(* CODESYS project filelogger.library
   DefaultNamespace: KOSTAL.AF2024.Core.FileLogger
   DocFormat: reStructuredText
   Description: Contains Functionalities to log strings to Filesystem with WSTRING content
   Author: Frank Dümpelmann
   Title: KOSTAL.AF2024.Core.FileLogger
   Version: 1.0.0.0
   Company: KOSTAL GmbH & Co.KG
   Placeholder: KOSTAL.AF2024.Core.FileLogger

Project tree, tasks and I/O mapping:
  libraries: KOSTAL.AF2024.Core.functionResponse, 1.0.0.0 (KOSTAL GmbH & Co.KG); KOSTAL.AF2024.Core.GetSystemTime, 1.0.0.0 (KOSTAL GmbH & Co.KG); KOSTAL.AF2024.Core.Process, 1.0.0.0 (KOSTAL GmbH & Co.KG); KOSTAL.AF2024.Core.Settings, 1.0.0.0 (KOSTAL GmbH & Co.KG); KOSTAL.AF2024.Core.StringTools, 1.0.0.0 (KOSTAL GmbH & Co.KG); KOSTAL.AF2024.Core.System, 1.0.0.0 (KOSTAL GmbH & Co.KG); Tc2_Standard, 3.3.3.0 (Beckhoff Automation GmbH); Tc2_System, 3.6.2.0 (Beckhoff Automation GmbH); Tc2_Utilities, 3.5.2.0 (Beckhoff Automation GmbH)
  DUT/
  POU/
    Interface/
      interface I_Logger: ePath, Extension, Path, Prefix, amsNedId_fileServer, delimiter, enabled, ID, maxLine, name, reset, StackCount, State, stepNumber, timeout, addLine
      interface I_Logger_Owner: ePath, Extension, Path, Prefix, amsNedId_fileServer, delimiter, enabled, maxLine, timeout, linkTimeSource, resetLogger, stepNumber
    function block FB_FileLogger [ST]: _a0_Ready, _a1_FileExist, _a2_Close, _a2_Open, _a2_Write, _Add_UTF16_LE_Header, _addLine, _control, _device, _formatWordToString, _getFqFileName, _outOfLimitControl, _stepHeader, _write, ePath, Extension, Path, Prefix, amsNedId_fileServer, delimiter, enabled, ID, maxLine, name, reset, StackCount, State, stepNumber, timeout, addLine, linkTimeSource, resetLogger, FBmain
  Project Information/
    function F_GetCompany [ST]
    function F_GetTitle [ST]
    function F_GetVersion [ST]
  Version/
    global variables Global_Version
*)

// Version/Global_Version
{attribute 'TcGenerated'}
{attribute 'no-analysis'}
{attribute 'linkalways'}
// This function has been automatically generated from the project information.
VAR_GLOBAL CONSTANT
	{attribute 'const_non_replaced'}
	stLibVersion_KOSTAL_AF2024_Core_FileLogger : ST_LibVersion := (iMajor := 1, iMinor := 0, iBuild := 0, iRevision := 0, nFlags := 0, sVersion := '1.0.0.0');
END_VAR

// POU/Interface/I_Logger
INTERFACE I_Logger EXTENDS KOSTAL_AF2024_Core_System.I_Interface

PROPERTY PUBLIC ePath : Tc2_System.E_OpenPath
GET
END_GET
END_PROPERTY

(*
Description
===========
| Extension of the saved file
| Default: .log
*)
PROPERTY PUBLIC Extension : STRING
GET
END_GET
END_PROPERTY

(*
Description
===========
| File path and name WITHOUT file extension
| e.g. "C:\\Logs\\test" creates the file "C:\\Logs\\test.log"
| default: c:\\temp\\log
*)
PROPERTY PUBLIC Path : KOSTAL_AF2024_Core_Settings.T_MaxString_UTF8
GET
END_GET
END_PROPERTY

PROPERTY PUBLIC Prefix : KOSTAL_AF2024_Core_Settings.T_MaxString_UTF8
GET
END_GET
END_PROPERTY

(*
Description
===========
| AMS NetID of  device to save log file to
| default: '' = Local device
*)
PROPERTY PUBLIC amsNedId_fileServer : STRING
GET
END_GET
END_PROPERTY

(*
Description
===========
| Delimiter to separate log records
| default: ;
*)
PROPERTY PUBLIC delimiter : WSTRING(1)
GET
END_GET
END_PROPERTY

(*
Description
===========
| Reset file handling sequence 
*)
PROPERTY PUBLIC enabled : BOOL
GET
END_GET
END_PROPERTY

PROPERTY ID : WSTRING
GET
END_GET
SET
END_SET
END_PROPERTY

(*
Description
===========
| Maximum number of message lines in write queue. 
| If the number is exceeded, the lines will be discarded
| default: 100, Maximum: 255
*)
PROPERTY PUBLIC maxLine : UDINT
GET
END_GET
END_PROPERTY

PROPERTY name : WSTRING
GET
END_GET
SET
END_SET
END_PROPERTY

(*
Description
===========
| Reset file handling sequence 
*)
PROPERTY PUBLIC reset : BOOL
GET
END_GET
END_PROPERTY

PROPERTY PUBLIC StackCount : UDINT
GET
END_GET
END_PROPERTY

PROPERTY PUBLIC State : KOSTAL_AF2024_Core_functionResponse.I_T_functionResponse
GET
END_GET
END_PROPERTY

PROPERTY stepNumber : INT
GET
END_GET
SET
END_SET
END_PROPERTY

(*
Description
===========
| Maximum time allowed for write operation
| default: 5s
*)
PROPERTY PUBLIC timeout : TIME
GET
END_GET
END_PROPERTY

(*
Description
===========
| Adds a line to the log file
| Parameters:
| 	line: KOSTAL_AF2024_Core_Settings.T_MaxString: Text to store in log file
| Return value:
| 	FB_functionResponse: 
|		result: BOOL: Operation succeeded
|		status: KOSTAL_AF2024_Core_Settings.T_MaxString:  Error description
*)

METHOD PUBLIC addLine : BOOL

VAR_INPUT
	line	: KOSTAL_AF2024_Core_Settings.T_MaxString;
END_VAR
END_METHOD

END_INTERFACE

// POU/Interface/I_Logger_Owner
INTERFACE I_Logger_Owner EXTENDS I_Logger

PROPERTY PUBLIC ePath : Tc2_System.E_OpenPath
SET
END_SET
END_PROPERTY

(*
Description
===========
| Extension of the saved file
| Default: .log
*)
PROPERTY PUBLIC Extension : STRING
SET
END_SET
END_PROPERTY

(*
Description
===========
| File path and name WITHOUT file extension
| e.g. "C:\\Logs\\test" creates the file "C:\\Logs\\test.log"
| default: c:\\temp\\log
*)
PROPERTY PUBLIC Path : KOSTAL_AF2024_Core_Settings.T_MaxString_UTF8
SET
END_SET
END_PROPERTY

PROPERTY PUBLIC Prefix : KOSTAL_AF2024_Core_Settings.T_MaxString_UTF8
SET
END_SET
END_PROPERTY

(*
Description
===========
| AMS NetID of  device to save log file to
| default: '' = Local device
*)
PROPERTY PUBLIC amsNedId_fileServer : STRING
SET
END_SET
END_PROPERTY

(*
Description
===========
| Delimiter to separate log records
| default: ;
*)
PROPERTY PUBLIC delimiter : WSTRING(1)
SET
END_SET
END_PROPERTY

(*
Description
===========
| Reset file handling sequence 
*)
PROPERTY PUBLIC enabled : BOOL
SET
END_SET
END_PROPERTY

(*
Description
===========
| Maximum number of message lines in write queue. 
| If the number is exceeded, the lines will be discarded
| default: 100, Maximum: 255
*)
PROPERTY PUBLIC maxLine : UDINT
SET
END_SET
END_PROPERTY

(*
Description
===========
| Maximum time allowed for write operation
| default: 5s
*)
PROPERTY PUBLIC timeout : TIME
SET
END_SET
END_PROPERTY

METHOD PUBLIC linkTimeSource
VAR_INPUT
	IN	: KOSTAL_AF2024_Core_GetSystemTime.I_TimeSource;
END_VAR
END_METHOD

METHOD PUBLIC resetLogger
VAR_INPUT
END_VAR
END_METHOD

PROPERTY stepNumber : INT
GET
END_GET
SET
END_SET
END_PROPERTY

END_INTERFACE

// POU/FB_FileLogger
(*

:Author: Frank Dümpelmann <f.duempelmann@kostal.com>
:Date: 2023-12-01

Function
========
Fuction block to write (WSTRING)lines to a log file in a specified location

Usage notes
===============
| Asyncronous function block: FB_Main() method must be called cyclicly
| Property getTimeStruct **must** be connected to a system time source, e.g. FB_get_NT_Clock
| Call Method addLine to write a string to the log file

Methods and Properties
======================
| See bottom of this document for a detailed description of each method or property
| Methods starting with an underline(_) are internally used and can be ignored by the user

Release Notes:
=============
| * V0.0.0.1

*)

FUNCTION_BLOCK PUBLIC FB_FileLogger IMPLEMENTS I_Logger_Owner, I_Logger

VAR
	_amsNedId_fileServer	: STRING:= '';	//default: local System
	_amsNedId_timeServer	: STRING:= '';	//default: local System
	
	{region 'file location'}
		_Path				: KOSTAL_AF2024_Core_Settings.T_MaxString_UTF8:= 'c:\temp\log\';	//default: 'c:\temp\log\'
		_Prefix			: KOSTAL_AF2024_Core_Settings.T_MaxString_UTF8:= 'log';	//default: log
		_Extension	: STRING:= 'log';	//default: 'log'
		_ePath			:	Tc2_System.E_OpenPath:= Tc2_System.E_OpenPath.PATH_GENERIC;	//default: PATH_GENERIC
	{endregion}
	
	_delimiter	: WSTRING(1)		:= ";";	//- default: "."

	_timeout	: TIME:= T#5S;	//- default: 5s
	
	_ID			: WSTRING;	//optional prefix after date and time in log line
	_name		: WSTRING;	//prefix after date and time in log line
	_stepNumber	: INT;

	_fileExist	: Tc2_Utilities.FB_EnumFindFileEntry;
	_fileDoExist: BOOL;
	
	_stack					: Kostal_AF2024_Core_StringTools.FB_ListOfString;
	_addLineContent			: KOSTAL_AF2024_Core_Settings.T_MaxString;	
	_line					: KOSTAL_AF2024_Core_Settings.T_MaxString; //stores the line input from addLine call
	
	_timeStamp	: KOSTAL_AF2024_Core_GetSystemTime.I_TimeSource;
	_openFile		: Tc2_System.FB_FileOpen;
	_writeFile	: Tc2_System.FB_FileWrite;
	_closeFile	: Tc2_System.FB_FileClose;

	_Step		: KOSTAL_AF2024_Core_process.FB_processStep_Flow;

	_writeLine	: KOSTAL_AF2024_Core_Settings.T_MaxString;	
	
	_enabled	: BOOL;	//BOOL
	_reset	: BOOL;
	_hFile	: UINT;

	_MonthAndYearForLog	: KOSTAL_AF2024_Core_Settings.T_MaxString;
	//_maxLine			: UDINT;

	
	_state	: KOSTAL_AF2024_Core_functionResponse.T_functionResponse;
	
END_VAR


VAR CONSTANT
	_ADDRESS_READY	: INT:= 0;
	_ADDRESS_CLOSE	: INT:= 3;
END_VAR

METHOD PROTECTED _a0_Ready
IF _Step.toggle THEN
	_closeFile.bExecute	:= FALSE;
	_openFile.bExecute	:= FALSE;
	_writeFile.bExecute	:= FALSE;
END_IF

_state.success	:= TRUE;
_state.status		:= "";

IF _Step.toggle THEN

	;	//do nothing

ELSIF _hFile <>  0 THEN

	_Step.set(_ADDRESS_CLOSE);
	
ELSIF  _stack.NumberOfLines = 0 THEN 

	_state.success	:= TRUE;
	_state.status		:= "stack is empty";

ELSE

	_state.success	:= TRUE;
	_state.status		:= "write line";


	_writeLine:= _stack.line_GET(1);
	_stack.removeLine(1);
	
	_Step.INC();
	
END_IF
END_METHOD

METHOD PROTECTED _a1_FileExist

IF _Step.toggle THEN
	_fileExist(bExecute:= TRUE, eCmd:= Tc2_Utilities.E_EnumCmdType.eEnumCmd_Abort);
	_fileExist(bExecute:= FALSE, eCmd:= Tc2_Utilities.E_EnumCmdType.eEnumCmd_Abort);
	_fileExist(bExecute:= TRUE, eCmd:= Tc2_Utilities.E_EnumCmdType.eEnumCmd_First, sPathName:= _getFqFileName());
END_IF

_fileExist(bExecute:= FALSE, eCmd:= Tc2_Utilities.E_EnumCmdType.eEnumCmd_First);

IF _fileExist.bBusy THEN

	_state.success:= TRUE;
	_state.status:= "try find file";

ELSIF _fileExist.bError THEN
	
	_state.success:= FALSE;
	_state.status:= Tc2_Standard.WCONCAT("Error find file with err.No.: ", UDINT_TO_WSTRING(_fileExist.nErrID)) ;
	
ELSE
	
	_fileDoExist:= _fileExist.stFindFile.sFileName <> '';

	_fileExist(bExecute:= TRUE, eCmd:= Tc2_Utilities.E_EnumCmdType.eEnumCmd_Abort);
	_fileExist(bExecute:= FALSE, eCmd:= Tc2_Utilities.E_EnumCmdType.eEnumCmd_Abort);

	_Step.INC();
	
END_IF
END_METHOD

METHOD PROTECTED _a2_Close
VAR_INPUT
END_VAR
IF _Step.toggle THEN
	_closeFile.bExecute:= FALSE;
END_IF

_state.success	:= TRUE;
_state.status		:= "";

IF _Step.toggle THEN

	_state.success	:= TRUE;
	_state.status		:= "close File - Init";

ELSIF NOT _closeFile.bExecute THEN

	_closeFile.bExecute:= TRUE;

	_state.success	:= TRUE;
	_state.status		:= "close File - Execute";

ELSIF _closeFile.bBusy THEN

	_state.success	:= TRUE;
	_state.status		:= "close File - Busy";


ELSIF _closeFile.bError THEN

	_state.success	:= FALSE;
	_state.status		:=  Tc2_Standard.WCONCAT("Error during close File. Err.ID > ", UDINT_TO_WSTRING(_closeFile.nErrId));
	
ELSE

	_state.success	:= TRUE;
	_state.status		:= "close File - Successful";

	_hFile:= 0;
	_Step.set(_ADDRESS_READY);
	
END_IF
END_METHOD

METHOD PROTECTED _a2_Open

IF _Step.toggle THEN
	
	_openFile.bExecute	:= FALSE;
	_openFile.sPathName:= _getFqFileName();
	
END_IF

_state.success	:= TRUE;
_state.status		:= "";

IF _Step.toggle THEN
	
	_state.success	:= TRUE;
	_state.status		:= "open File - Init";

ELSIF NOT _openFile.bExecute THEN

	_openFile.bExecute:= TRUE;

	_state.success	:= TRUE;
	_state.status		:= "open File - Execute";
	

ELSIF _openFile.bBusy THEN

	_state.success	:= TRUE;
	_state.status		:= "open File - Busy";

ELSIF _openFile.bError THEN

	_state.success	:= FALSE;
	_state.status		:=  Tc2_Standard.WCONCAT("Error during open File. Err.ID > ", UDINT_TO_WSTRING(_openFile.nErrId));
	
ELSE
	
	_hFile:= _openFile.hFile;
	
	_state.success	:= TRUE;
	_state.status		:= "open File - Successful";

	_Step.INC();
	
END_IF
END_METHOD

METHOD PROTECTED _a2_Write

VAR
	_concatLines	: ARRAY[1..14] OF KOSTAL_AF2024_Core_Settings.T_MaxString;
END_VAR


IF NOT _control() THEN RETURN;	END_IF

IF _Step.toggle THEN

	IF NOT _fileDoExist THEN _Add_UTF16_LE_Header();	END_IF

	_writeFile.bExecute	:= FALSE;

	_writeFile.pWriteBuff:= ADR(_writeLine);
	_writeFile.cbWriteLen:= INT_TO_UDINT((Tc2_Standard.WLEN(_writeLine) * 2) + 2);
	
END_IF


IF _Step.toggle THEN

	_state.success	:= TRUE;
	_state.status		:= "write File - Init";

ELSIF NOT _writeFile.bExecute THEN

	_writeFile.bExecute:= TRUE;

	_state.success	:= TRUE;
	_state.status		:= "write File - Execute";

ELSIF _writeFile.bBusy THEN

	_state.success	:= TRUE;
	_state.status		:= "write File - Busy";

ELSIF _writeFile.bError THEN

	_state.success	:= FALSE;
	_state.status		:=  Tc2_Standard.WCONCAT("Error during write File. Err.ID > ", UDINT_TO_WSTRING(_writeFile.nErrId));
	
ELSIF _stack.NumberOfLines > 0 THEN

	_state.success	:= TRUE;
	_state.status		:= "write line";

	_writeLine:= _stack.line_GET(1);
	_stack.removeLine(1);

	_writeFile.bExecute	:= FALSE;

	_writeFile.pWriteBuff:= ADR(_writeLine);
	_writeFile.cbWriteLen:= INT_TO_UDINT((Tc2_Standard.WLEN(_writeLine) * 2) + 2);

	
ELSE
	
	_state.success	:= TRUE;
	_state.status		:= "write File - Successful";
	
	_Step.INC();
	
END_IF
END_METHOD

METHOD PROTECTED _Add_UTF16_LE_Header

VAR
	_c: Kostal_AF2024_Core_StringTools.FB_Concat;
	_ws	: WSTRING;
	_p	: POINTER TO BYTE;
	
END_VAR

IF _p <> 0 THEN __DELETE(_p);	END_IF

_p:= __NEW(BYTE, (SIZEOF(_writeLine) + 2));

IF _p <> 0 THEN
	
	_p[0]:= 16#FF;
	_p[1]:= 16#FE;

	Tc2_System.MEMCPY((_p + 2), ADR(_writeLine), SIZEOF(_writeLine));

	_writeLine:= "";

	Tc2_System.MEMCPY(ADR(_writeLine), _p, SIZEOF(_writeLine));

	
END_IF
	
IF _p <> 0 THEN __DELETE(_p);	END_IF

(*
_p:= ADR(_ws);
_p[0]:= 16#FF;
_p[1]:= 16#FE;

_c.clear();
_c.addContent(_ws);
_c.addContent(_writeLine);

_writeLine:= _c.getResult();
_c.clear();
*)
END_METHOD

METHOD PROTECTED _addLine : BOOL

VAR
	_concat					:	Kostal_AF2024_Core_StringTools.FB_Concat;
END_VAR

_addLine:= FALSE;

IF _timeStamp = 0 										THEN _state.success:= FALSE;	_state.status:= "no (I_)Timestamp available";	RETURN;	END_IF
IF NOT _timeStamp.Valid	THEN _state.success:= FALSE;	_state.status:= "no valid Timestamp available";	RETURN;	END_IF

_concat.clear();
//Step  (optional)
//_concat.addContent(_addLineContent);

_concat.addContent(_name);
_concat.addContent(";");
_concat.addContent(INT_TO_WSTRING(_stepNumber));
_concat.addContent(";");

//_addLineContent:= _concat.getResult();

//ID (optional)
//_concat.clear();
//_concat.addContent(_addLineContent);

_concat.addContent(_ID);
_concat.addContent(";");

//_addLineContent:= _concat.getResult();

//Time
//_concat.clear();

//_concat.addContent(_addLineContent);
_concat.addContent(_formatWordToString(_timeStamp.timeStruct.Day, 2));
_concat.addContent(".");
_concat.addContent(_formatWordToString(_timeStamp.timeStruct.Month, 2));
_concat.addContent(".");
_concat.addContent( _formatWordToString(_timeStamp.timeStruct.Year, 4));

_concat.addContent(_delimiter);

_concat.addContent(_formatWordToString(_timeStamp.timeStruct.Hour, 2));
_concat.addContent(":");
_concat.addContent(_formatWordToString(_timeStamp.timeStruct.Minute, 2));
_concat.addContent(":");
_concat.addContent(_formatWordToString(_timeStamp.timeStruct.Second, 2));

_concat.addContent(_delimiter);

//Text
_concat.addContent(_line);

_concat.addContent("$R");

_addLineContent:= _concat.getResult();
_concat.clear();

_addLine:= TRUE;
END_METHOD

METHOD PROTECTED _control : BOOL
VAR_INPUT
END_VAR


_control:= FALSE;

IF _timeStamp = 0 THEN
	
	_state.status:= "getTimeStamp Reference is invalid";
	_state.success:= FALSE;

ELSIF NOT _timeStamp.Valid THEN
	
	_state.status:= "no valid timestamp available";
	_state.success:= FALSE;
	
ELSE

	_control:= TRUE;
	
	_state.status	:= "Control is successful";
	_state.success	:= TRUE;
	
END_IF
END_METHOD

METHOD PROTECTED _device

_fileExist(
	sNetId		:= _amsNedId_fileServer, 
	sPathName	:= , 
	eCmd			:= , 
	bExecute	:= , 
	tTimeout	:= _timeout, 
	bBusy				=> , 
	bError			=> , 
	nErrID			=> , 
	bEOE				=> , 
	stFindFile	=> );



_openFile
	(
		sNetId		:= _amsNedId_fileServer, 
		sPathName	:= , 
		nMode			:= Tc2_Utilities.FOPEN_MODEAPPEND, 
		ePath			:= _ePath, 
		bExecute	:= , 
		tTimeout	:= _timeout, 

		bBusy		=> , 
		bError	=> , 
		nErrId	=> , 
		hFile		=>	 
);

	_writeFile(
	sNetId			:= _amsNedId_fileServer, 
	hFile				:= _hFile, 
	pWriteBuff	:= , 
	cbWriteLen	:= , 
	bExecute		:= , 
	tTimeout		:= _timeout, 
	bBusy		=> , 
	bError	=> , 
	nErrId	=> , 
	cbWrite	=> );
	
_closeFile
	(
		sNetId		:= _amsNedId_fileServer, 
		hFile			:= _hFile, 
		bExecute	:= , 
		tTimeout	:= _timeout, 

		bBusy	=> , 
		bError=> , 
		nErrId=> 
	);
END_METHOD

METHOD PROTECTED _formatWordToString : KOSTAL_AF2024_Core_Settings.T_MaxString
VAR_INPUT
	IN			: WORD;
	length	: UINT;
END_VAR

_formatWordToString:= Tc2_Standard.WRIGHT(Tc2_Standard.WCONCAT("0000", WORD_TO_WSTRING(IN)), UINT_TO_INT(length));
END_METHOD

METHOD PROTECTED _getFqFileName : KOSTAL_AF2024_Core_Settings.T_MaxString_UTF8

VAR
	_c	: Kostal_AF2024_Core_StringTools.FB_Concat_UTF8;
	_pFix	: KOSTAL_AF2024_Core_Settings.T_MaxString_UTF8;
END_VAR

_c.Clear();

_c.addContent(_Path);

IF Tc2_Standard.RIGHT(_Path, 1) <> '\' THEN _c.addContent('\');	END_IF
	
IF _Prefix <> '' THEN _c.addContent(_Prefix);	_c.addContent('_');	END_IF

_c.addContent(WORD_TO_STRING(_timeStamp.timeStruct.Year));
_c.addContent('_');
_c.addContent(WORD_TO_STRING(_timeStamp.timeStruct.Month));

IF _Extension <> '' THEN
	IF Tc2_Standard.LEFT(_Extension, 1) <> '.' THEN	_c.addContent('.');	END_IF	
	_c.addContent(_Extension);
END_IF

_getFqFileName:= _c.getResult();

_c.Clear();
END_METHOD

METHOD PROTECTED _outOfLimitControl : BOOL
VAR_INPUT
END_VAR

IF _stack.NumberOfLines >= _stack.maxLine	THEN

	_outOfLimitControl := TRUE;
	_state.success:= FALSE;	
	_state.status:= "_outOfLimitControl - maxlines reached";	

END_IF
END_METHOD

METHOD PROTECTED _stepHeader
VAR_INPUT
END_VAR


IF _reset AND (_Step.actual > 0) THEN
	_Step.init();
 END_IF

_reset:= FALSE;

_Step.Header();
END_METHOD

METHOD PROTECTED _write


_stepHeader();

IF _Step.isActive(0)	THEN	_a0_Ready();			END_IF
IF _Step.isActive(1)	THEN	_a1_FileExist();	END_IF
IF _Step.isActive(2)	THEN	_a2_Open();				END_IF
IF _Step.isActive(3)	THEN	_a2_Write();			END_IF
IF _Step.isActive(4)	THEN	_a2_Close();			END_IF

IF _Step.NotFound()	THEN	
	_state.status		:= Tc2_Standard.WCONCAT("Step do not exist > ", INT_TO_WSTRING(_Step.actual));
	_state.success	:= FALSE;
END_IF
END_METHOD

PROPERTY PUBLIC ePath : Tc2_System.E_OpenPath
GET

ePath:= _ePath;
END_GET
SET

_ePath:= ePath;
END_SET
END_PROPERTY

(*
Description
===========
| Extension of the saved file
| Default: .log
*)
PROPERTY PUBLIC Extension : STRING
GET

Extension:= _Extension;
END_GET
SET

_Extension:= Extension;
END_SET
END_PROPERTY

(*
Description
===========
| File path and name WITHOUT file extension
| e.g. "C:\\Logs\\test" creates the file "C:\\Logs\\test.log"
| default: c:\\temp\\log
*)
PROPERTY PUBLIC Path : KOSTAL_AF2024_Core_Settings.T_MaxString_UTF8
GET

Path:= _Path;
END_GET
SET

_Path:= Path;
END_SET
END_PROPERTY

PROPERTY PUBLIC Prefix : KOSTAL_AF2024_Core_Settings.T_MaxString_UTF8
GET

Prefix:= _Prefix;
END_GET
SET

_Prefix:= Prefix;
END_SET
END_PROPERTY

(*
Description
===========
| AMS NetID of  device to save log file to
| default: '' = Local device
*)
PROPERTY PUBLIC amsNedId_fileServer : STRING
GET

amsNedId_fileServer:= _amsNedId_fileServer;
END_GET
SET

_amsNedId_fileServer:= amsNedId_fileServer;
END_SET
END_PROPERTY

(*
Description
===========
| Delimiter to separate log records
| default: ;
*)
PROPERTY PUBLIC delimiter : WSTRING(1)
GET

delimiter:= _delimiter;
END_GET
SET

_delimiter:= delimiter;
END_SET
END_PROPERTY

(*
Description
===========
| Reset file handling sequence 
*)
PROPERTY PUBLIC enabled : BOOL
GET

enabled:= _enabled;
END_GET
SET


_enabled:= enabled;
END_SET
END_PROPERTY

PROPERTY ID : WSTRING
GET

_ID:= _ID;
END_GET
SET

_ID:= ID;
END_SET
END_PROPERTY

(*
Description
===========
| Maximum number of message lines in write queue. 
| If the number is exceeded, the lines will be discarded
| default: 100, Maximum: 255
*)
PROPERTY PUBLIC maxLine : UDINT
GET

maxLine:= _stack.maxLine;
END_GET
SET


_stack.maxLine:= maxLine;
END_SET
END_PROPERTY

PROPERTY name : WSTRING
GET

name:= _name;
END_GET
SET

_name:= name;
END_SET
END_PROPERTY

(*
Description
===========
| Reset file handling sequence 
*)
PROPERTY PUBLIC reset : BOOL
GET

reset:= _reset;
END_GET
END_PROPERTY

PROPERTY PUBLIC StackCount : UDINT
GET

StackCount:= _stack.NumberOfLines;
END_GET
END_PROPERTY

PROPERTY PUBLIC State : KOSTAL_AF2024_Core_functionResponse.I_T_functionResponse
GET

state:= _state;
END_GET
END_PROPERTY

PROPERTY stepNumber : INT
GET

stepNumber:= _stepNumber;
END_GET
SET

_stepNumber:= stepNumber;
END_SET
END_PROPERTY

(*
Description
===========
| Maximum time allowed for write operation
| default: 5s
*)
PROPERTY PUBLIC timeout : TIME
GET

timeout:= _timeout;
END_GET
SET

_timeout:= timeout;
END_SET
END_PROPERTY

METHOD addLine : BOOL

VAR_INPUT
	line	: KOSTAL_AF2024_Core_Settings.T_MaxString;
END_VAR

IF NOT _enabled 				THEN RETURN;	END_IF
IF NOT _control() 			THEN RETURN;	END_IF
IF _outOfLimitControl()	THEN RETURN;	END_IF

_line:= line;
_addLineContent:= "";

addLine:= _addLine();

IF NOT addLine THEN RETURN;	END_IF

addLine:= _stack.addLine(_addLineContent);
END_METHOD

METHOD PUBLIC linkTimeSource
VAR_INPUT
	IN	: KOSTAL_AF2024_Core_GetSystemTime.I_TimeSource;
END_VAR

_timeStamp:= IN;
END_METHOD

METHOD PUBLIC resetLogger
VAR_INPUT
END_VAR

_reset:= TRUE;
END_METHOD

(*
Description
===========
| Main method, to be called cyclicly, e.g. in DeviceDefine
*)
METHOD PUBLIC FBmain

IF NOT _enabled THEN
	_state.status:= "not enabled";
	_state.success:= FALSE;
	RETURN;
END_IF

IF NOT _control() THEN RETURN;	END_IF

_device();

_write();
END_METHOD

END_FUNCTION_BLOCK

// Project Information/F_GetCompany
// This function has been automatically generated from the project information.
{attribute 'signature_flag' := '1073741824'}
{attribute 'TcGenerated'}
{attribute 'no-analysis'}
FUNCTION F_GetCompany : WSTRING
VAR_INPUT
	
END_VAR

F_GetCompany := "KOSTAL GmbH & Co.KG";

END_FUNCTION

// Project Information/F_GetTitle
// This function has been automatically generated from the project information.
{attribute 'signature_flag' := '1073741824'}
{attribute 'TcGenerated'}
{attribute 'no-analysis'}
FUNCTION F_GetTitle : WSTRING
VAR_INPUT
	
END_VAR

F_GetTitle := "KOSTAL.AF2024.Core.FileLogger";

END_FUNCTION

// Project Information/F_GetVersion
// This function has been automatically generated from the project information.
{attribute 'signature_flag' := '1073741824'}
{attribute 'TcGenerated'}
{attribute 'no-analysis'}
FUNCTION F_GetVersion : ST_LibVersion
VAR_INPUT
	
END_VAR

F_GetVersion.iMajor := 1;
F_GetVersion.iMinor := 0;
F_GetVersion.iBuild := 0;
F_GetVersion.iRevision := 0;
F_GetVersion.sVersion := '1.0.0.0';
F_GetVersion.nFlags := 0;

END_FUNCTION
